Fanuc KAREL source: kd00037.KL

-- PROVISIONAL review KL for V770-1; original PC SHA256 a5809ca2c7021476e32118359597f107e5de98e39f065b0b2d7d832cb575fa9a
-- Incomplete behavior may be omitted. Consult companion uncertainty JSON. Do not deploy.
PROGRAM KD00037
%NOLOCKGROUP
VAR
  I : INTEGER
  J : INTEGER
  B : BOOLEAN
  R : REAL
  S : STRING[80]
BEGIN
  -- UNRESOLVED_PC offsets 5-18; opcodes 9D,81,18,9D,1B,9D,12,9C,13,04
  -- UNRESOLVED_PC offsets 23-27; opcodes 7F
END KD00037
